{region 'Documentation'}
(*!
<summary>Checks equality with the expected BYTE value.</summary>
*)
{endregion}
FUNCTION_BLOCK AssertEqual_Byte EXTENDS AssertionBase
VAR_INPUT
    IN : BYTE; //! Actual value checked or observed by this Assertion.
    Expected : BYTE; //! Reference value for comparison with IN.
END_VAR

SUPER^();

{region 'Documentation'}
(*!
<summary>Check equality with the expected BYTE value.</summary>
*)
{endregion}
METHOD PROTECTED Assert
VAR
    Message : STRING(GVL_Constants.MessageLength);
    ExpectedText : STRING(GVL_Constants.AssertionValueLength);
    ActualText : STRING(GVL_Constants.AssertionValueLength);
END_VAR
VAR CONSTANT
    HexDigitCount : USINT := 2;
END_VAR
IF NOT EvaluationActive THEN
    RETURN;
END_IF;

IF Result = E_Result.Error THEN
    RETURN;
END_IF;

IF Result = E_Result.Failed THEN
    RETURN;
END_IF;

IF IN <> Expected THEN
    ExpectedText := CreateAssertionTextValue_Hex(Value := BYTE_TO_LWORD(Expected),
        DigitCount := HexDigitCount);
    ActualText := CreateAssertionTextValue_Hex(Value := BYTE_TO_LWORD(IN),
        DigitCount := HexDigitCount);
    Message := CONCAT('Assertion failed: values are not equal. Expected = ',
        ExpectedText);
    Message := CONCAT(Message, ', Actual = ');
    Message := CONCAT(Message, ActualText);
    Message := CONCAT(Message, '.');
    Fail(Message := Message);
    RETURN;
END_IF;

Pass();
END_METHOD

END_FUNCTION_BLOCK

(* stored: Version 1.1.0.1
   POU AssertEqual_Byte: Id {4bad0270-f7f0-42d6-b50f-de7b97b4f95e}, SpecialFunc None
   Folder Internal: Id {864824a7-9b90-4ec3-aee8-bb747dde3d25}
   Method Assert: Id {eae69aee-f50c-40be-a9a2-5c91c4706640} *)
